(* IEC 61131-3 sources: JingjiangArm/moonboxpro_arm_8.4/Application/Application/任务列表/TensionTask/电机运动, 6 files *)

(* ---- ENUM_AXISTYPE.st ---- *)
(*@CES
Name=ENUM_AXISTYPE
Type=Gvl
TypeGuid=2db5746d-d284-4425-9f7f-2663a34b0ebc
Guid=3491d2c6-312e-4e3b-a260-e28b79963db4
HasDeclaration=True
HasImplementation=False
*)
{DECLARATION}
TYPE ENUM_AXISTYPE :
(
	TYPE_MASTER_I,(*虚拟主轴/A系*)
	TYPE_MASTER_II,(*虚拟主轴/A系*)
	TYPE_CENTRAL_I,(*中心辊A*)
	TYPE_CENTRAL_II,(*中心辊B*)
	TYPE_UNWIND_A_I,(*放料A-A系*)
	TYPE_UNWIND_A_II,(*放料A-B系*)
	TYPE_UNWIND_B_I,(*放料B-A系*)
	TYPE_UNWIND_B_II,(*放料B-B系*)
	TYPE_REWIND_A_I,(*收料A-A系*)
	TYPE_REWIND_A_II,(*收料A-B系*)
	TYPE_REWIND_B_I,(*收料B-A系*)
	TYPE_REWIND_B_II,(*收料B-B系*)
	TYPE_INFEED_I,(*放牵A系*)
	TYPE_INFEED_II,(*放牵B系*)
	TYPE_OUTFEED_I,(*收牵A系*)
	TYPE_OUTFEED_II,(*收牵B系*)
	//TYPE_UNIT_CTL,(*色组控制轴@2026.5.20.135909 by liu.yt*)
	TYPE_UNIT_PRN,(*色组版辊*)
	TYPE_UNIT_ADJ,(*色组调整轴*)
	TYPE_UNIT_BOTTOM,(*色组底辊*)
	TYPE_UNIT_NET,(*色组网辊*)
	TYPE_UNIT_PRN_PRESS_MASTER,(*色组版辊龙门主轴*)
	TYPE_UNIT_PRN_PRESS_M,(*色组版辊龙门从轴M侧*)
	TYPE_UNIT_PRN_PRESS_G,(*色组版辊龙门从轴G侧*)
	TYPE_UNIT_NET_PRESS_MASTER,(*色组网辊龙门主轴*)
	TYPE_UNIT_NET_PRESS_M,(*色组网辊龙门从轴M侧*)
	TYPE_UNIT_NET_PRESS_G,(*色组网辊龙门从轴G侧*)
	TYPE_UNIT_STR_PRESS_MASTER,(*色组张带辊龙门主轴*)
	TYPE_UNIT_STR_PRESS_M,(*色组张带龙门从轴M侧*)
	TYPE_UNIT_STR_PRESS_G,(*色组张带龙门从轴G侧*)
	TYPE_UNIT_HORIZ,(*色组横向电机*)
	TYPE_UNIT_CTL,(*色组控制轴@2026.5.20.135909 by liu.yt*)
	TYPE_NULL(*未知*)
);
END_TYPE

{IMPLEMENTATION}

(* ---- ENUM_ControlledObjType.st ---- *)
(*@CES
Name=ENUM_ControlledObjType
Type=Gvl
TypeGuid=2db5746d-d284-4425-9f7f-2663a34b0ebc
Guid=c8e054b6-804a-4d86-ae05-73109a0c00ab
HasDeclaration=True
HasImplementation=False
*)
{DECLARATION}
TYPE ENUM_ControlledObjType :
(
	OBJ_IS_MASTERAXIS,(*主轴*)
	OBJ_IS_UNDEFINED,
	OBJ_IS_UNWIND_A,(* 放卷A *)
	OBJ_IS_UNWIND_B,(* 放卷B *)
	OBJ_IS_REWIND_A,(* 收卷A *)
	OBJ_IS_REWIND_B,(* 收卷B *)
	OBJ_IS_INFEED,(* 放牵 *)
	OBJ_IS_OUTFEED,(* 收牵 *)
	OBJ_IS_BOTTOM_ROLLER,(* 色组底辊 *)
	OBJ_IS_PRN_ROLLER,(* 色组版辊 *)

	OBJ_IS_NET_ROLLER,(* 色组网辊 *)
	OBJ_IS_PRN_ROLLER_PRESSURE_M,(* 色组版辊压力M侧 *)
	OBJ_IS_PRN_ROLLER_PRESSURE_G,(* 色组版辊压力G侧 *)

	OBJ_IS_NET_ROLLER_PRESSURE_M,(* 色组网辊压力M侧 *)
	OBJ_IS_NET_ROLLER_PRESSURE_G,(* 色组网辊压力G侧 *)
	OBJ_IS_STR_ROLLER_PRESSURE_M,(* 色组张带辊压力M侧 *)
	OBJ_IS_STR_ROLLER_PRESSURE_G,(* 色组张带辊压力G侧 *)
	OBJ_IS_HORIZ_MOTION,(* 横向运动电机/2022.6.8.142000 *)
	OBJ_IS_CENTRAL_DRUM,(* 中心滚筒/2022.6.8.135513 *)
	OBJ_IS_PHOTOCELL(*光电眼行走机构 | 2024.04.01.092649*)

);
END_TYPE

{IMPLEMENTATION}

(* ---- ENUM_MOTIONCTLSTEP.st ---- *)
(*@CES
Name=ENUM_MOTIONCTLSTEP
Type=Gvl
TypeGuid=2db5746d-d284-4425-9f7f-2663a34b0ebc
Guid=536e8cb1-3b5c-4e89-bb92-6c3fefab2bb0
HasDeclaration=True
HasImplementation=False
*)
{DECLARATION}
TYPE ENUM_MOTIONCTLSTEP :
(
	MOTION_STEP_Nothing,
	MOTIONCTL_STEP_SETMOTIONMODE,(*设置运动模式*)
	MOTIONCTL_STEP_RESET,(*初始化核*)
	MOTIONCTL_STEP_LOADWATCH,(**)
	MOTIONCTL_STEP_LMTSOFF,(*清除位置偏差报警*)
	MOTIONCTL_STEP_ALARMOFF,(*清除报警*)
	MOTIONCTL_STEP_ZEROPOS,(*清位置*)
	MOTIONCTL_STEP_CLRSTS,
	MOTIONCTL_STEP_AXISON,//上伺服
	MOTIONCTL_STEP_AXISOFF,//下伺服
	MOTIONCTL_STEP_CHECKAXISON,//检查使能状态
	MOTIONCTL_STEP_SETMODEPRM,//配置运动模式
	MOTIONCTL_STEP_WRITEDATA,//大指令数据填充
	MOTIONCTL_STEP_SetModal0				,(*2017-09-11 09:14:16| 模态0*)
	MOTIONCTL_STEP_SyncAllModal0				,(*同步所有轴模态|*)
	MOTIONCTL_STEP_SetModal1					,(*2017-09-11 09:14:24| 模态1*)
	MOTIONCTL_STEP_SyncAllModal1				,(*同步所有轴模态|*)
	MOTIONCTL_STEP_WaitingModalChanged	,	(*等待模态切换0到1|*)
	MOTIONCTL_STEP_WRITEDATA_Run,//大指令数据填充
	MOTIONCTL_STEP_WRITEDATA_Preg,//大指令数据填充
	MOTIONCTL_STEP_WRITEDATA_Inch,//大指令数据填充
	//2026.4.27.220207
	MOTIONCTL_STEP_WRITEDATA_Jog

);
END_TYPE

{IMPLEMENTATION}

(* ---- MotionSts.st ---- *)
(*@CES
Name=MotionSts
Type=Gvl
TypeGuid=2db5746d-d284-4425-9f7f-2663a34b0ebc
Guid=68a6a4b2-1fc3-48f5-a182-0781e2089d35
HasDeclaration=True
HasImplementation=False
*)
{DECLARATION}
{attribute 'pack_mode' := '1'}
TYPE MotionSts :
STRUCT
	lrMotionsts					: LREAL;
	lrPos_Prf					: LREAL;
	lrPos_Enc					: LREAL;
	lrVel_Prf					: LREAL;
	lrVel_Enc					: LREAL;
//扩展后，总共8个变量一张表
	lrAcc_Prf					: LREAL;
	lrTorque					: LREAL;
	lrData3						: LREAL;
END_STRUCT
END_TYPE

{IMPLEMENTATION}

(* ---- StUnitCfg.st ---- *)
(*@CES
Name=StUnitCfg
Type=Gvl
TypeGuid=2db5746d-d284-4425-9f7f-2663a34b0ebc
Guid=7ee9ace1-2ace-4dfd-ae7f-638a47057af9
HasDeclaration=True
HasImplementation=False
*)
{DECLARATION}
{attribute 'pack_mode' := '1'}
TYPE StUnitCfg :
STRUCT
	iUnitId : INT;
	iStationId : INT;
	iCoreId : INT;
	iAxisId : INT;
	iProfileId : INT;
	iAdjProfileId : INT;

END_STRUCT
END_TYPE

(*
TYPE StAxisCfg :
STRUCT
	iUnitId : INT;
	iStationId : INT;
	iCoreId : INT;
	iAxisId : INT;
	iProfileId : INT;
	iAdjProfileId : INT;

END_STRUCT
END_TYPE

*)
{IMPLEMENTATION}

(* ---- KS_HY_GetAxisIdForMotByStation.st ---- *)
(*@CES
Name=KS_HY_GetAxisIdForMotByStation
Type=FunctionBlock
TypeGuid=6f9dac99-8de1-4efc-8465-68ac443b7d08
Guid=98e977ff-93c3-495b-bafe-fe457f0448cc
HasDeclaration=True
HasImplementation=True
*)
{DECLARATION}
FUNCTION KS_HY_GetAxisIdForMotByStation : BOOL
VAR_INPUT
	i_iStationId: INT;
	i_piAxisId: POINTER TO INT;
	i_piTypeId: POINTER TO INT;
	i_piUnitId: POINTER TO INT;
	i_piCoreId: POINTER TO INT;
	i_piGroupId : POINTER TO INT;
	i_piAdjAxisId : POINTER TO INT;
	i_pastStAxisIdListInf: POINTER TO ARRAY [1..128] OF StAxisIdListInf;
END_VAR
VAR
	iN: INT;
	xResult: BOOL;
END_VAR

{IMPLEMENTATION}
xResult:= FALSE;
IF i_piAxisId<>0 AND i_piTypeId<>0 AND i_piUnitId<>0 AND i_piCoreId<>0 AND i_pastStAxisIdListInf<>0 AND
	i_iStationId>=0 AND i_iStationId< MAX_STATION_NUM THEN
	FOR iN:=1 TO 128 BY 1 DO
		IF i_iStationId= i_pastStAxisIdListInf^[iN].iStdId THEN
			i_piAxisId^:= i_pastStAxisIdListInf^[iN].iAxisId;
			i_piTypeId^:= i_pastStAxisIdListInf^[iN].iTypeId;
			i_piUnitId^:= i_pastStAxisIdListInf^[iN].iUnitId;
			i_piCoreId^:= i_pastStAxisIdListInf^[iN].iCoreId;
			i_piGroupId^:= i_pastStAxisIdListInf^[iN].iGroupId;
			i_piAdjAxisId^:= i_pastStAxisIdListInf^[iN].iAdjAxisId;
			EXIT;
		END_IF
	END_FOR
END_IF
